(* IEC 61131-3 sources: verifaps-lib/iec-symbex/src/test/resources/edu/kit/iti/formal/automation/rvt, 4 files *)

(* ---- effective_subtypes.st ---- *)
INTERFACE ITF
  METHOD f : INT
    VAR_INPUT
      x : INT;
    END_VAR
  END_METHOD
END_INTERFACE

CLASS A IMPLEMENTS ITF
  VAR
    b1 : B;
    b2 : B;
    c1 : C;
    c2 : C;
  END_VAR

  METHOD f : INT
    VAR_INPUT
      x : INT;
    END_VAR

    b1.c1.z := FALSE;
    f := 42;
  END_METHOD
END_CLASS

CLASS A1 EXTENDS A
  METHOD f : INT
    VAR_INPUT
      x : INT;
    END_VAR

    f := 24;
  END_METHOD
END_CLASS

CLASS A2 EXTENDS A
  METHOD f : INT
    VAR_INPUT
      x : INT;
    END_VAR

    f := 33;
  END_METHOD
END_CLASS

CLASS B IMPLEMENTS ITF
  VAR
    c1 : C;
    c2 : C;
  END_VAR
END_CLASS

CLASS C
  VAR
    z : BOOL;
  END_VAR
END_CLASS

PROGRAM MY_PROGRAM
  VAR_INPUT
    switch : BOOL;
    x : INT;
  END_VAR
  VAR
    i : ITF;
    a : A;
    a1 : A1;
    b : B;
    r : REF_TO A;
  END_VAR
  VAR_OUTPUT
    y : INT;
  END_VAR

  r := REF(a1);

  IF (switch) THEN
    i := a;
  ELSE
    i := b;
  END_IF

  y := r^.f(x);

  r^.c1 := a.b1.c1;
  r^.c2 := a.b2.c2;

  r^.b1.c2 := r^.c2;
END_PROGRAM

(* ---- effective_subtypes_no_methods.st ---- *)
CLASS A
  VAR
    c1 : C;
    c2 : C;
  END_VAR
END_CLASS

CLASS A1 EXTENDS A
END_CLASS

CLASS A2 EXTENDS A
END_CLASS

CLASS C
  VAR
    z : INT;
  END_VAR
END_CLASS

PROGRAM MY_PROGRAM
  VAR_INPUT
    switch : BOOL;
    x : INT;
  END_VAR
  VAR
    a : A;
    a1 : A1;
    r : REF_TO A;
  END_VAR
  VAR_OUTPUT
    y : INT;
  END_VAR

  IF (switch) THEN
    r := REF(a);
  ELSE
    r := REF(a1);
  END_IF

  r^.c1.z := x;
  r^.c2.z := x + 2;

  IF (switch) THEN
    y := r^.c1.z;
  ELSE
    y := r^.c2.z;
  END_IF

  y := y + x;
END_PROGRAM

(* ---- references.st ---- *)
INTERFACE ITF1
  METHOD func : INT
  END_METHOD
END_INTERFACE

INTERFACE ITF2
END_INTERFACE

INTERFACE ITF3
END_INTERFACE

CLASS ClBase IMPLEMENTS ITF1, ITF2
  VAR
    x : INT;
  END_VAR

  METHOD func : INT
    func := 42;
  END_METHOD
END_CLASS

CLASS ClDerived EXTENDS ClBase IMPLEMENTS ITF3
  METHOD func : INT
    func := 24;
  END_METHOD
END_CLASS

PROGRAM MY_PROGRAM
  VAR
    instBase : ClBase;
    instDerived: ClDerived;
    rinstBase1, rinstBase2: REF_TO ClBase;
    rinstDerived1, rinstDerived2: REF_TO ClDerived;
    rinstDerived3, rinstDerived4: REF_TO ClDerived;
    interf1: ITF1;
    interf2: ITF2;
    interf3: ITF3;
  END_VAR

rinstBase1:= REF(instBase); // rinstbase1 references base class
rinstBase2:= REF(instDerived); // rinstbase2 references derived class

rinstDerived1 ?= rinstBase1; // rinstDerived1 == NULL
rinstDerived2 ?= rinstBase2; // rinstDerived2 will contain a valid
                             // reference to instDerived
interf1:= instBase;    // interf1 is a reference to base class
interf2:= instDerived; // interf2 is a reference to derived class

rinstDerived3 ?= interf1; // rinstDerived3 == NULL
rinstDerived4 ?= interf2; // rinstDerived4 will contain a valid
                          // reference to instDerived

rinstBase1:= REF(instBase); // rinstbase1 references base class
rinstBase2:= REF(instDerived); // rinstbase2 references derived class

rinstBase1^.x := interf1.func();  // 42
rinstBase2^.x := interf2.func();  // 24

END_PROGRAM

(* ---- simple_hierarchy.st ---- *)
CLASS A
  VAR
    x : INT;
    y : INT;
  END_VAR

  METHOD f : INT
    x := x + 1;
    f := x + y;
  END_METHOD

  METHOD g : INT
    y := y + 1;
    g := x * y;
  END_METHOD
END_CLASS

CLASS B EXTENDS A
  VAR
    z : INT;
  END_VAR

  METHOD OVERRIDE f : INT
    f := SUPER.f() + z;
  END_METHOD

  METHOD OVERRIDE g : INT
    z := z - 1;
    g := x * y * z;
  END_METHOD
END_CLASS

CLASS C EXTENDS B
  VAR
    r : INT;
  END_VAR

  METHOD OVERRIDE g : INT
    g := r * x * y * z;
  END_METHOD
END_CLASS

PROGRAM MY_PROGRAM
  VAR
    a : A := (x := 42, y := 24);
    b : B := (x := 33, y := 44, z := 55);
    c : C := (x := 1, y := 2, z := 3, r := 4);
  END_VAR
  VAR_OUTPUT
    x : INT;
    y : INT;
  END_VAR

  y := c.f();
  x := c.x;
END_PROGRAM
